FUNCTION_BLOCK IO_AO (* One analog output, also a PWM channel (the step pulses of a stepper motor, a motor's speed). Its Address says where it goes: a Raspberry Pi PWM channel, a Modbus register, or simulated. Technical: Analog output (raw = Bias + OUT * Gain, 0..65535; EN = FALSE writes 0); Address: 'gpio[chip:line(:pull_up|:pull_down)(:active_low)]' or 'pwm[chip:channel:period_ns]' a Raspberry Pi's line, set up here; 'modbus[...]' a Modbus CLIENT ID; 'sim' simulated; another name a local IO handle set up elsewhere (QW PARAMS); empty: not connected (QO = FALSE) *)
  (* Standard: 61499-2 *)
  (* Version 0.1, 2026-09-28, Project contributors, AAU Smart Production Lab *)
  PACKAGE modlib;
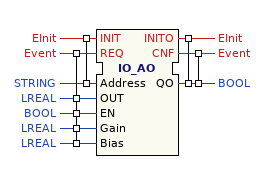
  EVENT_INPUT
    INIT : EInit WITH Address; (* Set up the point from Address (at start-up) *)
    REQ WITH OUT, EN, Gain, Bias; (* Read the point, or write OUT to it *)
  END_EVENT
  EVENT_OUTPUT
    INITO : EInit WITH QO; (* Set up: QO says whether the point is reachable *)
    CNF WITH QO; (* Done: QO says whether it worked (an input: IN is the value read) *)
  END_EVENT
  VAR_INPUT
    Address : STRING; (* Where the point is: 'gpio[chip:line(:pull_up|:pull_down)(:active_low)]', 'pwm[chip:channel:period_ns]', 'modbus[...]', 'sim', or an IO handle's name; empty: not connected *)
    OUT : LREAL; (* The value to write *)
    EN : BOOL; (* On; FALSE writes 0 (no pulses on a PWM channel) *)
    Gain : LREAL := 1.0; (* Raw = Bias + OUT * Gain, limited to 0..65535 *)
    Bias : LREAL; (* Raw = Bias + OUT * Gain, limited to 0..65535 *)
  END_VAR
  VAR_OUTPUT
    QO : BOOL; (* The point is reachable, the last access worked *)
  END_VAR
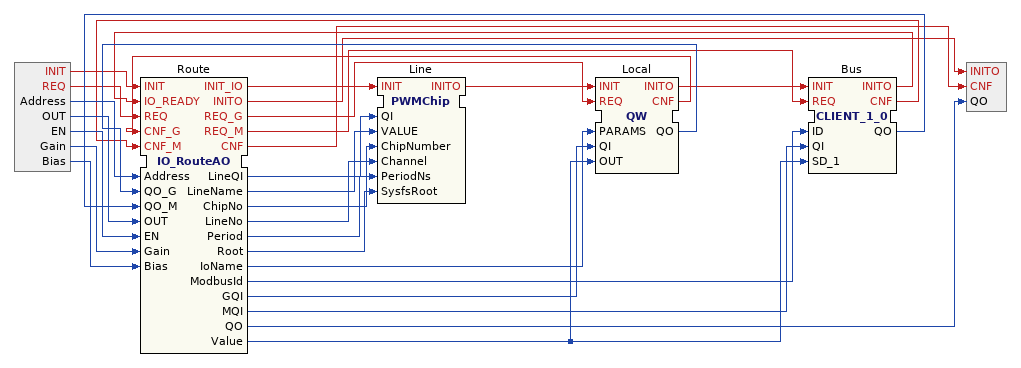
  FBS
    Route : modlib::IO_RouteAO; (* Picks the way to the signal from the Address and passes values that way. *)
    Line : eclipse4diac::io::pwmsysfs::PWMChip; (* Sets up a Raspberry Pi line (GPIO) or PWM channel when the Address names one. *)
    Local : eclipse4diac::io::QW; (* Reads or writes a FORTE IO handle (IX, QX, IW, QW). *)
    Bus : iec61499::net::CLIENT_1_0; (* Reads or writes a Modbus register when the Address names one. *)
  END_FBS
  EVENT_CONNECTIONS
    INIT TO Route.INIT;
    Route.INIT_IO TO Line.INIT;
    Line.INITO TO Local.INIT;
    Local.INITO TO Bus.INIT;
    Bus.INITO TO Route.IO_READY;
    Route.INITO TO INITO;
    REQ TO Route.REQ;
    Route.REQ_G TO Local.REQ;
    Route.REQ_M TO Bus.REQ;
    Local.CNF TO Route.CNF_G;
    Bus.CNF TO Route.CNF_M;
    Route.CNF TO CNF;
  END_CONNECTIONS
  DATA_CONNECTIONS
    Route.LineQI TO Line.QI;
    Route.LineName TO Line.VALUE;
    Route.ChipNo TO Line.ChipNumber;
    Route.LineNo TO Line.Channel;
    Route.Period TO Line.PeriodNs;
    Route.Root TO Line.SysfsRoot;
    Address TO Route.Address;
    Route.IoName TO Local.PARAMS;
    Route.ModbusId TO Bus.ID;
    Route.GQI TO Local.QI;
    Route.MQI TO Bus.QI;
    Local.QO TO Route.QO_G;
    Bus.QO TO Route.QO_M;
    Route.QO TO QO;
    OUT TO Route.OUT;
    EN TO Route.EN;
    Gain TO Route.Gain;
    Bias TO Route.Bias;
    Route.Value TO Local.OUT;
    Route.Value TO Bus.SD_1;
  END_CONNECTIONS
END_FUNCTION_BLOCK
